FUNCTION F_OpcUaCreateSubscribeId (* Creates an OPC UA identifier for a subscription *)
  (* Standard: 61499-2; Description: Copyright (c) 2026 Monika Wenger This program and the accompanying materials are made available under the terms of the Eclipse Public License 2.0 which is available at https://www.eclipse.org/legal/epl-2.0/ SPDX-License-Identifier: EPL-2.0 *)
  (* Version 3.0, 2026-10-14, Monika Wenger *)
  PACKAGE eclipse4diac::opcua;
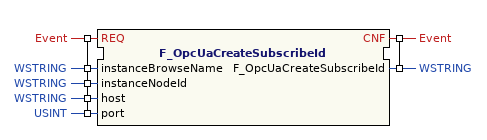
  EVENT_INPUT
    REQ WITH instanceBrowseName, instanceNodeId, host, port;
  END_EVENT
  EVENT_OUTPUT
    CNF WITH F_OpcUaCreateSubscribeId;
  END_EVENT
  VAR_INPUT
    instanceBrowseName : WSTRING;
    instanceNodeId : WSTRING;
    host : WSTRING;
    port : USINT;
  END_VAR
  VAR_OUTPUT
    F_OpcUaCreateSubscribeId : WSTRING;
  END_VAR
  BODY IN ST:
PACKAGE eclipse4diac::opcua;

(* Creates an OPC UA identifier for a subscription *)
FUNCTION F_OpcUaCreateSubscribeId : WSTRING
VAR_INPUT
	instanceBrowseName : WSTRING;
	instanceNodeId : WSTRING;
	host : WSTRING;
	port : USINT;
END_VAR
VAR CONSTANT
	PREFIX : WSTRING := "opc_ua[SUBSCRIBE;opc.tcp://";
	NODEID_TYPE : WSTRING := ",s=";
	SUFFIX : WSTRING := "]";
	SEPARATOR_HASH : WSTRING := "#;";
	SEPARATOR_HOST : WSTRING := ":";
END_VAR
F_OpcUaCreateSubscribeId := CONCAT(PREFIX, host, SEPARATOR_HOST, USINT_AS_WSTRING(port), SEPARATOR_HASH,
	instanceBrowseName, NODEID_TYPE, instanceNodeId, SUFFIX);
END_FUNCTION
  END_BODY
END_FUNCTION
